// TIA Portal V21 export
// export: Created 2026-08-21T20:18:57.0934095Z, ExportSetting None, DisplayName Totally Integrated Automation Portal, DisplayVersion V21, DisplayName STEP 7 Professional, DisplayVersion V21, DisplayName STEP 7 Safety, DisplayVersion V21, DisplayName Tech WebApplication, DisplayVersion V21, DisplayName WinCC Basic/Comfort/Advanced, DisplayVersion V21, DisplayName WinCC Professional, DisplayVersion V21, DisplayName WinCC Unified, DisplayVersion V21
TYPE "UDT_Service_Value"
   STRUCT
      Analog : Real;   // Analog value
      Digital : DInt;   // Digital value
      Binary : Bool;   // Binary value
      "String" : String[40];   // String value
   END_STRUCT;
END_TYPE
